TYPE ST_PNOZData :
STRUCT
    //Project identification
    wsProjectName: WSTRING(16);
    nProjectChecksum: WORD;
    nOverallChecksum: WORD;

    //Project creation date
    sCreationDate: STRING(10); //E.g. 2026.3.4


    //Additional stored date and time
    sStoredDate: STRING(18); //E.g. 2026.11.12 44h 13m

    //Operating-hours snapshot
    nOperatingHoursAtInit: UDINT;

    //Modules
    stBaseUnit: ST_PNOZModuleData;
    stFieldbus: ST_PNOZModuleData;

    astRightModule: ARRAY[1..MAX(USINT#1, GVL_APP.nNUM_OF_EXPANSION_RIGHT)] OF ST_PNOZModuleData;
    astLeftModule: ARRAY[1..MAX(USINT#1, GVL_APP.nNUM_OF_EXPANSION_LEFT)] OF ST_PNOZModuleData;
END_STRUCT
END_TYPE

(* stored: Version 1.1.0.1
   DUT ST_PNOZData: Id {edbe01c0-bb8e-07e4-0dc0-7cf94a8e0c1a} *)
